Fanuc KAREL source: KD00044.KL

PROGRAM KD00044
%NOLOCKGROUP
VAR
  I: INTEGER
  J: INTEGER
  B: BOOLEAN
  R: REAL
  S: STRING[80]
  G: GROUP_ASSOC
BEGIN
  I = 1
END KD00044
